(* PLC project g_star_delta_no_deadtime, Anonymous Benchmark Suite 1.0 *)
(* stored: creationDateTime 2026-08-28T00:00:00 *)

PROGRAM g_star_delta_no_deadtime
  VAR_INPUT
    Call : BOOL;
    StarDone : BOOL;
    DeadDone : BOOL;
  END_VAR
  VAR_OUTPUT
    Star : BOOL;
    Delta : BOOL;
  END_VAR

(* LD diagram, written out as Structured Text *)
Star := Call AND NOT StarDone;
Delta := Call AND StarDone;
END_PROGRAM

CONFIGURATION Config0
  RESOURCE Res0 ON PLC
    TASK tcyclic(INTERVAL := T#10ms, PRIORITY := 0);
    PROGRAM inst0 WITH tcyclic : g_star_delta_no_deadtime;
  END_RESOURCE
END_CONFIGURATION
